// TIA Portal V20 export
TYPE "WT3_Verdichter_Status_UDT"
   STRUCT
      iHandshake : Int;
      Alarm : Struct
         bE0000_KonfigAlarm : Bool;
         bE0001_VerbundMasterAusg : Bool;
         bE0002_NotstoppPHDFehler : Bool;
         bE0003_ExternAlarm : Bool;
         bE0004_TDruckAlarm : Bool;
         bE0005_PDruckAlarm : Bool;
         bE0006_PSaugAlarm : Bool;
         bE0007_TMotorAlarm : Bool;
         bE0008_TSHMinSaugAlarm : Bool;
         bE0009_TSHMinDruckAlarm : Bool;
         bE0010_LuefterAlarm : Bool;
         bE0011_Reserviert : Bool;
         bE0012_PhasenFehler : Bool;
         bE0013_MotorAlarm : Bool;
         bE0014_LSAusloesung : Bool;
         bE0015_POeldiffStillstand : Bool;
         bE0016_POeldiffBetrieb : Bool;
         bE0017_TOelMaxAlarm : Bool;
         bE0018_OElniveauOA : Bool;
         bE0019_OElniveauVd : Bool;
         bE0020_OElStroemung : Bool;
         bE0021_POelfilterBetrieb : Bool;
         bE0022_TLagerDEAlarm : Bool;
         bE0023_TLager_NDEAlarm : Bool;
         bE0024_Reserviert : Bool;
         bE0025_Reserviert : Bool;
         bE0026_Reserviert : Bool;
         bE0027_PSaugOverrange : Bool;
         bE0028_PPsZuTief : Bool;
         bE0029_Oelpumpe : Bool;
         bE0030_Leistungsschieber : Bool;
         bE0031_PoPsZuTief : Bool;
         bE0032_StartdruckZuHoch : Bool;
         bE0033_POelfilterStillstand : Bool;
         bE0034_PoPMinAlarm : Bool;
         bE0035_Startoeldruck : Bool;
         bE0036_TDruckGradient : Bool;
         bE0037_OelflussVerdichter : Bool;
         bE0038_KeineGasfoerderung : Bool;
         bE0039_PZwDruck : Bool;
         bE0040_TZwDruck : Bool;
         bE0041_TSHMinZwDruck : Bool;
         bE0042_POeldiffMax : Bool;
         bE0043_PPsMax : Bool;
         bE0044_OelkhlungTop : Bool;
         bE0045_PPzZuTeif : Bool;
         bE0046_PPzMax : Bool;
         bE0047_PPsZuTief : Bool;
         bE0048_FluessigSchlag : Bool;
         bE0049_Reserviert : Bool;
         bE0050_Reserviert : Bool;
         bE0051_Reserviert : Bool;
         bE0052_Reserviert : Bool;
         bE0053_Reserviert : Bool;
         bE0054_Reserviert : Bool;
         bE0055_Reserviert : Bool;
         bE0056_Reserviert : Bool;
         bE0057_Reserviert : Bool;
         bE0058_Reserviert : Bool;
         bE0059_Reserviert : Bool;
         bE0060_Reserviert : Bool;
         bE0061_Reserviert : Bool;
         bE0062_Reserviert : Bool;
         bE0063_KaeltekreisMasterAusgefa : Bool;
         bE0064_Reserviert : Bool;
         bE0065_KaelteKreisInvUngueltig : Bool;
         bE0066_OelkreisMasterAusgefa : Bool;
         bE0067_Reserviert : Bool;
         bE0068_OelKreisInvUngueltig : Bool;
         bE0069_SchmierdruckMin : Bool;
         bE0070_PPoMax : Bool;
         bE0071_Haupt_OeldruckMin : Bool;
         bE0072_Reserviert : Bool;
         bE0073_Reserviert : Bool;
         bE0074_Reserviert : Bool;
         bE0075_TZylinderkopfAlarm : Bool;
         bE0076_VerdampferpumpeAlarmBet : Bool;
         bE0077_VerdampferpumpeAlarmSti : Bool;
         bE0078_NivHDAbschHochAlarm : Bool;
         bE0079_NivEconomiserHochAlarm : Bool;
         bE0080_Reserviert : Bool;
         bE0081_KonfAlarmKkStart_Stopp : Bool;
         bE0082_HDVerdAusgefallen : Bool;
         bE0083_NDVerdAusgefallen : Bool;
         bE0084_KeinStartbefehlKonf : Bool;
         bE0085_PzPsMax : Bool;
         bE0086_Reserviert : Bool;
         bE0087_VibraSwitchAusg : Bool;
         bE0088_TOelabschMax : Bool;
         bE0089_TOelMin : Bool;
         bE0090_Reserviert : Bool;
         bE0091_NDAbschNivHoch : Bool;
         bE0092_Sekundaerschieber : Bool;
         bE0093_Reserviert : Bool;
         bE0094_KonfigAlarmAbsKuehls : Bool;
         bE0095_Reserviert : Bool;
         bE0096_OelnivKGHhoch : Bool;
         bE0097_KonfigAlarmDIPrio : Bool;
         bE0098_Reserviert : Bool;
         bE0099_Reserviert : Bool;
         bE0100_Reserviert : Bool;
         bE0101_KonfigAlarmDrehzahl : Bool;
         bE0102_Reserviert : Bool;
         bE0103_PSaugHoch : Bool;
         bE0104_KonfigAlarmMotorleist : Bool;
         bE0105_AlarmEinsatzdiagr : Bool;
         bE0106_Reserviert : Bool;
         bE0107_Reserviert : Bool;
         bE0108_Reserviert : Bool;
         bE0109_MotorAlarmNotAusTest : Bool;
         bE0110_StirnspHauptrotorZGross : Bool;
         bE0111_StirnspHautprotorZKlein : Bool;
         bE0112_StirnspNebenrotorZGross : Bool;
         bE0113_StirnspNebenrotorZKlein : Bool;
         bE0114_THauptrotorDS : Bool;
         bE0115_THauptrotorSS : Bool;
         bE0116_TNebenrotorDS : Bool;
         bE0117_TNebenrotorSS : Bool;
         bE0118_FlSchlagAlarmSensor : Bool;
         bE0119_OelstoppventilAlarm : Bool;
         bE0120_Reserviert : Bool;
         bE0121_Reserviert : Bool;
         bE0122_Reserviert : Bool;
         bE0123_Reserviert : Bool;
         bE0124_Reserviert : Bool;
         bE0125_Reserviert : Bool;
         bE0126_Reserviert : Bool;
         bE0127_Reserviert : Bool;
         bE0128_Reserviert : Bool;
         bE0129_Reserviert : Bool;
         bE0130_Reserviert : Bool;
         bE0131_Reserviert : Bool;
         bE0132_Reserviert : Bool;
         bE0133_Reserviert : Bool;
         bE0134_Reserviert : Bool;
         bE0135_Reserviert : Bool;
         bE0136_Reserviert : Bool;
         bE0137_Reserviert : Bool;
         bE0138_VorschmierenNötig : Bool;
         bE0139_KonfigAlarmHltebetrieb : Bool;
         bE0140_AlarmTTOPHKZuTief : Bool;
         bE0141_AlarmTTOPHKZuHoch : Bool;
         bE0142_KonfigAlarmKeinDefVi : Bool;
         bE0143_Reserviert : Bool;
         bE0144_Reserviert : Bool;
         bE0145_ÖlabscheiderStartniveauTief : Bool;
         bE0146_Reserviert : Bool;
         bE0147_PSaugGradientHochFehler : Bool;
         bE0148_UEGAlarm : Bool;
         bE0149_TechStrömungGMA : Bool;
         bE0150_VerdichterAutomatikbetriebNichtMöglich : Bool;
         bE0151_FuStörung : Bool;
         b210_Reserve : Bool;
         bE0153_RevSchalterVerdichterMotorImBetrieb : Bool;
         bE0154_KonfigFehlerFuStartdrehzahl : Bool;
         bE0155_AlarmStartdrehzahlNichtErreicht : Bool;
         bE0156_AlarmFuStartzeitZuKurz : Bool;
         b215_Reserve : Bool;
         bE0158_SammelstörungSchieberansteuerung : Bool;
         bE0159_RevisionsschalterÖlpumpe : Bool;
         "bE0160_Alarm PDruckseitePÖlausgleichskolben" : Bool;
         bE0161_AlarmPDruckseitePInjektionöl : Bool;
         bE0162_NothaltSR1PZhFehler : Bool;
         bE0163_AbsperrhahnDruckseiteNichtOffen : Bool;
         bE0164_AbsperrhahnDruckseiteNichtZu : Bool;
         bE0165_AbsperrhahnSaugseiteNichtOffen : Bool;
         bE0166_AbsperrhahnSaugseiteNichtZu : Bool;
         bE0167_Reserviert : Bool;
         bE0168_AbsperrhahnEconomiserNichtOffen : Bool;
         bE0169_AbsperrhahnEconomiserNichtZu : Bool;
         bE0170_Reserviert : Bool;
         bE0171_SpeisungMagnetventile230V : Bool;
         "bE0172_AlarmP-Öldifferenzschwingt" : Bool;
         bE0173_StartvorhaltZuLange : Bool;
         "bE0174_VSE135_S1.1_Alarm" : Bool;
         "bE0175_VSE135_S1.2_Alarm" : Bool;
         "bE0176_VSE135_S2.1_Alarm" : Bool;
         "bE0177_VSE135_S2.2_Alarm" : Bool;
         "bE0178_VSE135_S3.1_Alarm" : Bool;
         "bE0179_VSE135_S3.2_Alarm" : Bool;
         "bE0180_VSE135_S3.4_Alarm" : Bool;
         "bE0181_VSE135_S4.1_Alarm" : Bool;
         "bE0182_VSE135_S4.2_Alarm" : Bool;
         "bE0183_VSE135_S4.3_Alarm" : Bool;
         "bE0184_VSE135_S4.4_Alarm" : Bool;
         "bE0185_VSE135_S4.5_Alarm" : Bool;
         b252_Reserve : Bool;
         b253_Reserve : Bool;
         bE0188_StörungÜberhitzungsventil : Bool;
         bE0189_SoftstarterStörung : Bool;
         bE0190_StörungEconomiserventil : Bool;
         bE0200_AlarmKabelbruch : Bool;
         by26_Reserve : Byte;
         by27_Reserve : Byte;
         by28_Reserve : Byte;
         by29_Reserve : Byte;
         by30_Reserve : Byte;
         by31_Reserve : Byte;
         by32_Reserve : Byte;
         by33_Reserve : Byte;
      END_STRUCT;
      Warnung : Struct
         bA1000_Reserviert : Bool;
         bA1001_VerbundMasterAusg : Bool;
         bA1002_Reserviert : Bool;
         bA1003_Reserviert : Bool;
         bA1004_TDruck : Bool;
         bA1005_PDruck : Bool;
         bA1006_Reserviert : Bool;
         bA1007_TMotor : Bool;
         bA1008_TSHMinSaug : Bool;
         bA1009_TSHMinDruck : Bool;
         bA1010_Reserviert : Bool;
         bA1011_Reserviert : Bool;
         bA1012_Reserviert : Bool;
         bA1013_Reserviert : Bool;
         bA1014_Reserviert : Bool;
         bA1015_Reserviert : Bool;
         bA1016_POeldiff_Betrieb : Bool;
         bA1017_TOelmax : Bool;
         bA1018_OelniveauOA : Bool;
         bA1019_Reserviert : Bool;
         bA1020_Reserviert : Bool;
         bA1021_POelfilterBetrieb : Bool;
         bA1022_TLagerDE : Bool;
         bA1023_TLagerNDE : Bool;
         bA1024_OelniveauOA_hoch : Bool;
         bA1025_Reserviert : Bool;
         bA1026_Reserviert : Bool;
         bA1027_PSaugOverrange : Bool;
         bA1028_PPszutief : Bool;
         bA1029_Reserviert : Bool;
         bA1030_Reserviert : Bool;
         bA1031_Reserviert : Bool;
         bA1032_Reserviert : Bool;
         bA1033_Reserviert : Bool;
         bA1034_PoPMin : Bool;
         bA1035_Reserviert : Bool;
         bA1036_Reserviert : Bool;
         bA1037_Reserviert : Bool;
         bA1038_Reserviert : Bool;
         bA1039_PZwDruck : Bool;
         bA1040_TZwDruck : Bool;
         bA1041_TSHminZwDruck : Bool;
         bA1042_Reserviert : Bool;
         bA1043_PPsmax : Bool;
         bA1044_Reserviert : Bool;
         bA1045_PPzzutief : Bool;
         bA1046_PPzmax : Bool;
         bA1047_PPszutief2 : Bool;
         bA1048_FluessigSchlag : Bool;
         bA1049_NDPendel : Bool;
         bA1050_TOelMin : Bool;
         bA1051_Reserviert : Bool;
         bA1052_OelheizungOA : Bool;
         bA1053_TSaug : Bool;
         bA1054_PSauglimit : Bool;
         bA1055_PDrucklimit : Bool;
         bA1056_LastabwurfMotorstrom : Bool;
         bA1057_MinLeistungnErr : Bool;
         bA1058_MaxLeistungnErr : Bool;
         bA1059_BalanceFNorm : Bool;
         bA1060_PrimaerschMaxNErr : Bool;
         bA1061_LastabwurfMotorleistung : Bool;
         bA1062_OelheizungKGH : Bool;
         bA1063_KaeltekreisMasterAusgef : Bool;
         bA1064_KaeltekreisSlaveAusgef : Bool;
         bA1065_Reserviert : Bool;
         bA1066_Reserviert : Bool;
         bA1067_OelkreisSlaveAusgef : Bool;
         bA1068_Reserviert : Bool;
         bA1069_SchmierdruckMin : Bool;
         bA1070_PPoMax : Bool;
         bA1071_HauptOeldruckMin : Bool;
         bA1072_Oelnachspeisung : Bool;
         bA1073_KdMasterAusgef : Bool;
         bA1074_VrMasterAusgef : Bool;
         bA1075_TZylinderkopf : Bool;
         bA1076_Reserviert : Bool;
         bA1077_Reserviert : Bool;
         bA1078_Reserviert : Bool;
         bA1079_Reserviert : Bool;
         bA1080_KdMasterAusef : Bool;
         bA1081_Reserviert : Bool;
         bA1082_Reserviert : Bool;
         bA1083_Reserviert : Bool;
         bA1084_Reserviert : Bool;
         bA1085_PzPsWarnung : Bool;
         bA1086_HauptMasterAusgef : Bool;
         bA1087_Reserviert : Bool;
         bA1088_TOelabschMaxWarnung : Bool;
         bA1089_TOelMinWarnung : Bool;
         bA1090_OelpumpePendelwarnung : Bool;
         bA1091_Reserviert : Bool;
         bA1092_Reserviert : Bool;
         bA1093_TOelMinWarnungKGH : Bool;
         bA1094_Reserviert : Bool;
         bA1095_TZwDruckSaugHDWarnung : Bool;
         bA1096_OelniveauKGHHoch : Bool;
         bA1097_Reserviert : Bool;
         bA1098_MKaeltekrMasterAktiv : Bool;
         bA1099_MOelkreisMasterAktiv : Bool;
         "bA1100_Objekt-ID mehrfach vorhanden" : Bool;
         bA1101_Reserviert : Bool;
         bA1102_RekalibrierungMinNDurchg : Bool;
         bA1103_Reserviert : Bool;
         bA1104_Reserviert : Bool;
         bA1105_WarnungEinsatzdiagr : Bool;
         bA1106_WarnungEcoNivEndsch : Bool;
         bA1107_OelnachspDVrGesp : Bool;
         bA1108_OerektDVrGesp : Bool;
         bA1109_NotAusTestFehlgeschl : Bool;
         bA1110_StirnspHauptrotorZGross : Bool;
         bA1111_StirnspHauptrotorZKlein : Bool;
         bA1112_StirnspNebenrotorZGross : Bool;
         bA1113_StirnspNebenrotorZKlein : Bool;
         bA1114_THauptrotorDS : Bool;
         bA1115_THauptrotorSS : Bool;
         bA1116_TNebenrotorDS : Bool;
         bA1117_TNebenrotorSS : Bool;
         bA1118_FlSchlagWarnungSensor : Bool;
         bA1119_Reserviert : Bool;
         bA1120_PDruckMinWarnung : Bool;
         bA1121_Vorschm10Tagen : Bool;
         bA1122_Vorschm9Tagen : Bool;
         bA1123_Vorschm8Tagen : Bool;
         bA1124_Vorschm7Tagen : Bool;
         bA1125_Vorschm6Tagen : Bool;
         bA1126_Vorschm5Tagen : Bool;
         bA1127_Vorschm4Tagen : Bool;
         bA1128_Vorschm3Tagen : Bool;
         bA1129_Vorschm2Tagen : Bool;
         bA1130_Vorschm1Tag : Bool;
         bA1131_Reserviert : Bool;
         bA1132_Reserviert : Bool;
         bA1133_Reserviert : Bool;
         bA1134_Reserviert : Bool;
         bA1135_Reserviert : Bool;
         bA1136_Reserviert : Bool;
         bA1137_Reserviert : Bool;
         bA1138_Reserviert : Bool;
         bA1139_Reserviert : Bool;
         bA1140_WarnungTTOPHKZuTief : Bool;
         bA1141_WarnungTTOPHKZuHoch : Bool;
         bA1142_Reserviert : Bool;
         bA1143_PlusSperreDruckseite : Bool;
         bA1144_PlusSperreSaugseite : Bool;
         bA1145_Reserviert : Bool;
         bA1146_DruckabfallFeinabscheider : Bool;
         bA1147_PSaugGradientHochWarnung : Bool;
         bA1148_Reserviert : Bool;
         bA1149_Reserviert : Bool;
         b526_Reserve : Bool;
         b527_Reserve : Bool;
         bA1152_StrömungswächterWHC : Bool;
         b531_Reserve : Bool;
         b532_Reserve : Bool;
         bA1155_AlarmStartdrehzahlNichtErreicht : Bool;
         bA1156_AlarmFUStartzeitZuKurz : Bool;
         bA1157_ExternFreigabeÖlnaschspFehlt : Bool;
         b536_Reserve : Bool;
         b537_Reserve : Bool;
         bA1160_bAlarmPDruckseitePÖlausgleichskolben : Bool;
         bA1161_bAlarmPDruckseitePInjektionöl : Bool;
         bA1162_Reserviert : Bool;
         bA1163_Reserviert : Bool;
         bA1164_Reserviert : Bool;
         bA1165_Reserviert : Bool;
         bA1166_Reserviert : Bool;
         bA1167_SchieberStartpositionNichtErreicht : Bool;
         bA1168_Reserviert : Bool;
         bA1169_Reserviert : Bool;
         bA1170_StartdruckZuTief : Bool;
         bA1171_Reserviert : Bool;
         "bA1172_WarnungP-ÖldifferenzSchwingt" : Bool;
         bA1173_Reserviert : Bool;
         "bA1174_VSE135_S1.1_Warnung" : Bool;
         "bA1175_VSE135_S1.2_Warnung" : Bool;
         "bA1176_VSE135_S2.1_Warnung" : Bool;
         "bA1177_VSE135_S2.2_Warnung" : Bool;
         "bA1178_VSE135_S3.1_Warnung" : Bool;
         "bA1179_VSE135_S3.2_Warnung" : Bool;
         "bA1180_VSE135_S3.4_Warnung" : Bool;
         "bA1181_VSE135_S4.1_Warnung" : Bool;
         "bA1182_VSE135_S4.2_Warnung" : Bool;
         "bA1183_VSE135_S4.3_Warnung" : Bool;
         "bA1184_VSE135_S4.4_Warnung" : Bool;
         "bA1185_VSE135_S4.5_Warnung" : Bool;
         bA1186_WarnungVSE135Kommunikation : Bool;
         bA1187_SensorfehlerVibrationsmessgerät : Bool;
         bA1188_Reserviert : Bool;
         bA1189_Reserviert : Bool;
         bA1190_Reserviert : Bool;
         bA1191_Reserviert : Bool;
         by58_Reserve : Byte;
         bA1200_WarnungKabelbruch : Bool;
         b591_Reserve : Bool;
         b592_Reserve : Bool;
         b593_Reserve : Bool;
         b594_Reserve : Bool;
         b595_Reserve : Bool;
         b596_Reserve : Bool;
         b597_Reserve : Bool;
         by60_Reserve : Byte;
         by61_Reserve : Byte;
         by62_Reserve : Byte;
         by63_Reserve : Byte;
         by64_Reserve : Byte;
         by65_Reserve : Byte;
      END_STRUCT;
      Zustand : Struct
         bAlarmzustandAktiv : Bool;
         bWarnzustandAktiv : Bool;
         bSystemMeldungAktiv : Bool;
         bServiceMeldungAktiv : Bool;
         bStopManuell : Bool;
         bStopAuto : Bool;
         bStopExtern : Bool;
         bBetriebAuto : Bool;
         bBetriebManuell : Bool;
         bAnlaufAuto : Bool;
         bAnlaufManuell : Bool;
         bManuellStoppen : Bool;
         b674_Reserve : Bool;
         b675_Reserve : Bool;
         b676_Reserve : Bool;
         b677_Reserve : Bool;
         by68_Reserve : Byte;
         by69_Reserve : Byte;
         bAnlaufsperre : Bool;
         bVerdichterSaugtAb : Bool;
         bLastabwurfSaugseite : Bool;
         bLastabwurfDruckseite : Bool;
         bLastabwurfPPs : Bool;
         bElStromGrNormal : Bool;
         bElStromGrMaximum : Bool;
         bOelZuKalt : Bool;
         bNiveauOelabschZuTief : Bool;
         bExternsperreAktiv : Bool;
         b712_Reserviert : Bool;
         b713_Reserviert : Bool;
         bExternLimitAktiv : Bool;
         bInternLimitAktiv : Bool;
         bVerdichterVollOel : Bool;
         b717_Reserviert : Bool;
         b720_Reserviert : Bool;
         bSealLube : Bool;
         bKeineFrgZwischendruck : Bool;
         bElLeistungGrNormal : Bool;
         bElLeistungGrMaximum : Bool;
         bBegrElLeistungAkt : Bool;
         bStartbefehlManuell : Bool;
         bOelpumpeManuell : Bool;
         bOelrektifizierungMan : Bool;
         bOelkuehlerManuell : Bool;
         bInventarKaeltekreis : Bool;
         bInventarOelkreis : Bool;
         bMasterGesperrt : Bool;
         bKaeltekrStbyMstInit : Bool;
         bKaeltekrStbyMstPassiv : Bool;
         bKaeltekrStbyMstAktiv : Bool;
         bHaltManuell : Bool;
         bGesperrtVonKd : Bool;
         bGesperrtVonVr : Bool;
         bOelZuWarm : Bool;
         bNachkalMin : Bool;
         bPDruckZuHoch : Bool;
         bVdStartVerz : Bool;
         bSchieberZwangstr : Bool;
         bGespVonOelkreisMaster : Bool;
         PDruckLimitAktiv : Bool;
         PDruckGradLimitAktiv : Bool;
         PSaugLimitAktiv : Bool;
         PSaugGradLimitAktiv : Bool;
         "bSchmierungN.Stillstand" : Bool;
         bÖlabscheiderLimitAktiv : Bool;
         "bSperreTopH/K" : Bool;
         PlusSperreDruckseite : Bool;
         PlusSperreSaugseite : Bool;
         bGenerellGesperrt : Bool;
         b763_Reserve : Bool;
         bFUNichtBereit : Bool;
         bAbsperrventileWerdenGeöffnet : Bool;
         "bFU-RampeAktiv" : Bool;
         bSoftstarterNichtBereit : Bool;
         bGesperrtDurchKältekreis : Bool;
         "bGesperrtDurchVr-Pumpe" : Bool;
         "bGesperrtDurchKd-Pumpe" : Bool;
         b773_Reserve : Bool;
         b774_Reserve : Bool;
         b775_Reserve : Bool;
         b776_Reserve : Bool;
         b777_Reserve : Bool;
         by78_Reserve : Byte;
         by79_Reserve : Byte;
         by80_Reserve : Byte;
         by81_Reserve : Byte;
      END_STRUCT;
      "Allgemeine Meldungen" : Struct
         b4000_AllgemeineMeldung_1 : Bool;
         b4001_AllgemeineMeldung_2 : Bool;
         b4002_AllgemeineMeldung_3 : Bool;
         b4003_AllgemeineMeldung_4 : Bool;
         b4004_AllgemeineMeldung_5 : Bool;
         b4005_AllgemeineMeldung_6 : Bool;
         b4006_AllgemeineMeldung_7 : Bool;
         b4007_AllgemeineMeldung_8 : Bool;
         by83_Reserve : Byte;
         by84_Reserve : Byte;
         by85_Reserve : Byte;
      END_STRUCT;
      DigIn : Struct
         bNotstopp : Bool;
         bFehlerExtern : Bool;
         bPhasenuberwachung : Bool;
         bNiveauOelabscheiderTief : Bool;
         bNiveauOelabscheiderHoch : Bool;
         bNiveauKurbelgehaeuseTief : Bool;
         b866_Reserviert : Bool;
         bStartbefehl : Bool;
         bRmVerdichtermotor : Bool;
         bRmElOelpumpe : Bool;
         bExternLeistungslimit : Bool;
         bStartprioritaet : Bool;
         bRmChillerpumpe : Bool;
         b875_Reserviert : Bool;
         bMotorbegrenzung : Bool;
         bPDruckseiteDigital : Bool;
         bPSaugseiteDigital : Bool;
         bPOelLubeDigital : Bool;
         bPOelfilterDigital : Bool;
         bTDruckseiteDigital : Bool;
         b884_Reserviert : Bool;
         bTOelDigital : Bool;
         bTOelabscheiderDigital : Bool;
         bTMotorDigital : Bool;
         bNivKurbelGehaeuseHoch : Bool;
         bRueckmeldungLuefter : Bool;
         bRueckmeldungStoerung : Bool;
         bNivNDAbschHoch : Bool;
         bNivEconomiserHoch : Bool;
         bLastsperre : Bool;
         b896_Reserviert : Bool;
         bOelstrBitzer : Bool;
         bOelflussYork : Bool;
         bOelabschNivNormal : Bool;
         bAuxDigital1 : Bool;
         bAuxDigital2 : Bool;
         bVerdichterOelniveau : Bool;
         bVibraSwitch : Bool;
         bNDAbschNiveauHochMax : Bool;
         bStartzwangExtern : Bool;
         bOelnivKurbelGehaeuseNorm : Bool;
         bExternsperre : Bool;
         bDrehmomentbegrenzung : Bool;
         bNiveauEconomOpen : Bool;
         bNiveauEconomClose : Bool;
         bOelstoppventilBitzer : Bool;
         bFreigabePDruckLimit : Bool;
         bFreigabePSaugLimit : Bool;
         bFreigabeHaltebetrieb : Bool;
         bSperreGenerell : Bool;
         bAlarmUEG : Bool;
         BTechnischeStörungGMA : Bool;
         bFUStörung : Bool;
         bVdMotorRevSchalter : Bool;
         bFUBereit : Bool;
         bStrömungswächterWHC : Bool;
         bÖlnachspeisungExtFreigabe : Bool;
         bSammelstörungSchiebersteuerung : Bool;
         bRevisionsschalterÖlpumpe : Bool;
         bNothaltSicherheitsrelais1 : Bool;
         bEndschalterAbsperrhahnDruckseiteOffen : Bool;
         bEndschalterAbsperrhahnSaugseiteOffen : Bool;
         bEndschalterAbsperrhahnDruckseiteZu : Bool;
         bEndschalterAbsperrhahnSaugseiteZu : Bool;
         bDrehzahlbegrenzungTief : Bool;
         bDrehzahlbegrenzungHoch : Bool;
         bLeistungMinErhöhen : Bool;
         bAbsperrhahnEcoOffen : Bool;
         bAbsperrhahnEcoZu : Bool;
         b945_Reserve : Bool;
         b946_Reserve : Bool;
         b947_Reserve : Bool;
         by95_Reserve : Byte;
         by96_Reserve : Byte;
         by97_Reserve : Byte;
         by98_Reserve : Byte;
         by99_Reserve : Byte;
         by100_Reserve : Byte;
         by101_Reserve : Byte;
      END_STRUCT;
      DigOut : Struct
         bAlarm : Bool;
         bWarnung : Bool;
         bLastschalterAusloesung : Bool;
         bBereit : Bool;
         bStart_Motor : Bool;
         bAnlaufentlastung : Bool;
         bTeilwicklung2 : Bool;
         bMagnetventilFluessig : Bool;
         bOelheizungOelabscheider : Bool;
         bOelheizungKurbelgehaeuse : Bool;
         bStartOelpumpe : Bool;
         bOelventil : Bool;
         bOelrektifizierungA : Bool;
         bOelrektifizierungB : Bool;
         bOelrueckfuehrung : Bool;
         bOelnachspeisung : Bool;
         bOelkuehlung : Bool;
         bPowerkit : Bool;
         bEconomiser : Bool;
         bLeistungGrGrenzwert : Bool;
         bZwischendruckkuehlung : Bool;
         bVerdapferpumpe : Bool;
         bStartanzeige : Bool;
         bGrundlastzylinder : Bool;
         bViMax : Bool;
         bViMin : Bool;
         bVi22 : Bool;
         bVi2235 : Bool;
         bUeberhitzungsventil : Bool;
         bStillstandentlastung : Bool;
         bOeltransfer : Bool;
         bFastPullDownMV : Bool;
         bNiveaureglerEconom : Bool;
         bOelrektEinzeln : Bool;
         bSaugleitungsheizung : Bool;
         bLeistungsschPulsBitzer : Bool;
         bAnzSchmierungNStillstand : Bool;
         bTOPHeizung : Bool;
         bTOPMVKuehlen : Bool;
         bHauptÖlventil : Bool;
         bMVFlüssigInjektion : Bool;
         bQuittieranzeigeNothaltFehler : Bool;
         bQuittieranzeigeNothaltSR1Fehler : Bool;
         bQuittieranzeigeNothaltSR2Fehler : Bool;
         bQuittieranzeigeAlarmUEG : Bool;
         bQuittieranzeigeFUStörung : Bool;
         bStoppanzeige : Bool;
         bSchieberQuittierung : Bool;
         bSammelsignalWarnung : Bool;
         bSammelsignalAlarm : Bool;
         bResetFuSRSignal : Bool;
         bAbsperrhahnDruckseite : Bool;
         bAbsperrhahnSaugseite : Bool;
         bMVFlüssigkeitsableitungSaugleitung : Bool;
         bAbsperrhahnEconomiser : Bool;
         bLeistungsventil1 : Bool;
         bLeistungsventil2 : Bool;
         bLeistungsventil3 : Bool;
         bLeistungsventil4 : Bool;
         bLeistungsventil5 : Bool;
         bLeistungsventil6 : Bool;
         bLeistungsventil7 : Bool;
         b1096_Reserve : Bool;
         b1097_Reserve : Bool;
         by110_Reserve : Byte;
         by111_Reserve : Byte;
         by112_Reserve : Byte;
         by113_Reserve : Byte;
         by114_Reserve : Byte;
         by115_Reserve : Byte;
         by116_Reserve : Byte;
         by117_Reserve : Byte;
      END_STRUCT;
      rPDruckBar : Real;
      rPDruckGrad : Real;
      rPSaugBar : Real;
      rPSaugGrad : Real;
      rIstleistProz : Real;
      rIstleistVol : Real;
      rSollleistProz : Real;
      rSollleistVol : Real;
      rIstVi : Real;
      rSollVi : Real;
      rPZwStufeBar : Real;
      rPZwStufeGrad : Real;
      rPEcoBar : Real;
      rPEcoGrad : Real;
      rPOelLube : Real;
      rPOelDiff : Real;
      rPOelfilter : Real;
      rPOelpumpe : Real;
      rPKGH : Real;
      rTDruck : Real;
      rTSaug : Real;
      rTZwStufe : Real;
      rTOel : Real;
      rTOelabscheider : Real;
      rTSHDruck : Real;
      rTSHSaug : Real;
      rTSHZwStufe : Real;
      rMotorstromA : Real;
      rMotorstromProz : Real;
      rMotorleistkW : Real;
      rMotorleistProz : Real;
      rMotorPTC : Real;
      diEinschaltMotor : DInt;
      diBetriebsstunden : DInt;
      iAktVdStufe : Int;
      rOelkRegIst : Real;
      rOelkRegSoll : Real;
      rOelkRegOut : Real;
      rMotordrehzahl : Real;
      diEnergiezaehlerTot : DInt;
      rOaNiveau : Real;
      rAuxAnalog1 : Real;
      rMinLeistung : Real;
      rMaxLeistung : Real;
      rPOelfilterEinAus : Real;
      rTOelkuehlerEin : Real;
      rTOelkuehlerAus : Real;
      rPosPriSchieber : Real;
      rPosSekSchieber : Real;
      rTSaugleitung : Real;
      rNDAbscheiderNiveau : Real;
      rEconomiserNiveau : Real;
      rTVerdichterkühlAustritt : Real;
      rTZwStufeSaugHD : Real;
      rTEconomiser : Real;
      rTTOPHeizenKühlen : Real;
      rEconomiserAnalog : Real;
      rUeberhitzungsventil : Real;
      rAnlaufentlastungAnalog : Real;
      rOelpumpenAusgang : Real;
      rEcoNiveaureglerAusgang : Real;
      diLaeuftSeit : DInt;
      rCPos : Real;
      rFUIstfrequenz : Real;
      rFUSollwert : Real;
      rCabs : Real;
      rNullpositionSchieber : Real;
      diModus : DInt;
      rMotortemperaturU1 : Real;
      rMotortemperaturV1 : Real;
      rMotortemperaturW1 : Real;
      rMotortemperaturU2 : Real;
      rMotortemperaturV2 : Real;
      rMotortemperaturW2 : Real;
      rTMotorlagerDE : Real;
      rTMotorlagerNDE : Real;
      rPosPrimärschieberSoll : Real;
      rPosSekundärschieberSoll : Real;
      rTZylinderkopf1 : Real;
      rTZylinderkopf2 : Real;
      rTZylinderkopf3 : Real;
      rTZylinderkopf4 : Real;
      rTZylinderkopf5 : Real;
      rTZylinderkopf6 : Real;
      rTZylinderkopf7 : Real;
      rTZylinderkopf8 : Real;
      rTZylinderkopf9 : Real;
      rTZylinderkopf10 : Real;
      rTZylinderkopf11 : Real;
      rTZylinderkopf12 : Real;
      rTZylinderkopf13 : Real;
      rTZylinderkopf14 : Real;
      rTZylinderkopf15 : Real;
      rTZylinderkopf16 : Real;
      rPDruck_PSaug_Differenz : Real;
      rPDruck_PSaug_Verhältniss : Real;
      rPDruck_PZwStufe_Differenz : Real;
      rPDruck_PZwStufe_Verhältniss : Real;
      rPZwStufe_PSaug_Differenz : Real;
      rTHauptrotorlagerDS : Real;
      rTHauptrotorlagerSS : Real;
      rTNebenrotorlagerDS : Real;
      rTNebenrotorlagerSS : Real;
      diStufePreset : DInt;
      rPFeinabscheiderEintritt : Real;
      rPFeinabscheiderAustritt : Real;
      rGasKonzentration : Real;
      rPEco_PSaug_Differenz : Real;
      rStirnspaltHauptrotorDiff : Real;
      rStirnspaltHauptrotor : Real;
      rStirnspaltNebenrotorDiff : Real;
      rStirnspaltNebenrotor : Real;
      rMinVerflüssigungsTemperatur : Real;
      rFlüssInjection : Real;
      rÖlInjection : Real;
      rTSHDruckSoll : Real;
      rEnergiezählerTrip : Real;
      diVerdichterstartsHeute : DInt;
      diVerdichterstartsGestern : DInt;
      dikontrolleVerdichterLagerSeitService : DInt;
      diKontrolleVerdichterLagerBisService : DInt;
      diKontrolleMotorLagerSeitService : DInt;
      diKontrolleMotorLagerBisService : DInt;
      diKontrolleWellenabdichtungSeitService : DInt;
      diKontrolleWellenabdichtungBisService : DInt;
      diKontrolleSaugDruckVentileSeitService : DInt;
      diKontrolleSaugDruckVentileBisService : DInt;
      diKontrolleMotorschmierungSeitService : DInt;
      diKontrolleMotorschmierungbisService : DInt;
      diÖlanalyseSeitService : DInt;
      diÖlanalyseBisService : DInt;
      diÖltestSeitService : DInt;
      diÖltestBisService : DInt;
      diÖlwechselSeitService : DInt;
      diÖlwechselBisService : DInt;
      diLetzteDynWartungA : DInt;
      dinächsteDynWartungA : DInt;
      diLetzteDynWartungB : DInt;
      diNächsteDynWartungB : DInt;
      diLetzteDynWartungC : DInt;
      diNächsteDynWartungC : DInt;
      rAuxAnalog2 : Real;
      rPÖlausgleichskolben : Real;
      rPInjektionöl : Real;
      rDrehzahlbegrenzungTief : Real;
      rDrehzahlbegrenzungHoch : Real;
      rSchieberStellwert : Real;
      diPrioritätsstunden : DInt;
      rTOPDreiwegventilKühlen : Real;
      rBetriebsmodusAktiv : Real;
      byReserve : Array[716..1023] of Byte;
   END_STRUCT;
END_TYPE
